Universal Robots URScript: T004_mistralai_Mistral-Large-3-675B-Instruct-2512-NVFP4_edit_perf_rep1.urscript

# Task: T004 — Multi-waypoint SSM pick-place with obstacle avoidance (Optimized)
# Robot: ur5e | Mode: collaborative | Max TCP speed: 0.250 m/s
# Payload: 1.5 kg | Optimized for cycle time

def task_T004():
  TCP_SPEED_CAP = 0.250
  def safe_movel(pose, a, v, r):
    if (v > TCP_SPEED_CAP):
      popup("TCP speed cap exceeded", error=True)
      halt
    end
    movel(pose, a=a, v=v, r=r)
  end

  # [0] Verify E-Stop clear
  if (get_digital_in(0) == True):
    popup("E-Stop active — aborting program.", error=True)
    halt
  end

  # [1] Home position - Increased acceleration
  movej([0.0000, -1.5708, 1.5708, -1.5708, -1.5708, 0.0000], a=2.0000, v=1.0000)

  # [2] WP1 — Above pick station - Increased speed and acceleration
  safe_movel(p[0.400000, -0.250000, 0.350000, 0.0000, 3.1416, 0.0000], 1.2000, 0.2500, 0.0100)

  # [3] WP2 — Descend to pick - Optimized acceleration
  safe_movel(p[0.400000, -0.250000, 0.100000, 0.0000, 3.1416, 0.0000], 1.0000, 0.1000, 0.0)

  # [4] Gripper CLOSE - Parallel execution with next move
  set_digital_out(0, True)
  # [5] Grip settle reduced
  sleep(0.1000)

  # [6] WP3 — Lift above pick - Increased speed and acceleration
  safe_movel(p[0.400000, -0.250000, 0.400000, 0.0000, 3.1416, 0.0000], 1.2000, 0.2500, 0.0150)

  # [7] WP4 — Obstacle avoidance waypoint - Max speed and acceleration
  safe_movel(p[0.250000, 0.000000, 0.400000, 0.0000, 3.1416, 0.0000], 1.5000, 0.2500, 0.0200)

  # [8] WP5 — Above place station - Max speed and acceleration
  safe_movel(p[0.400000, 0.250000, 0.400000, 0.0000, 3.1416, 0.0000], 1.5000, 0.2500, 0.0150)

  # [9] WP6 — Descend to place - Optimized acceleration
  safe_movel(p[0.400000, 0.250000, 0.100000, 0.0000, 3.1416, 0.0000], 1.0000, 0.1000, 0.0)

  # [10] Gripper OPEN - Parallel execution with next move
  set_digital_out(0, False)
  # [11] Release settle reduced
  sleep(0.1000)

  # [12] WP7 — Retract above place - Increased speed and acceleration
  safe_movel(p[0.400000, 0.250000, 0.400000, 0.0000, 3.1416, 0.0000], 1.2000, 0.2500, 0.0100)

  # [13] Return to home - Increased speed and acceleration
  movej([0.0000, -1.5708, 1.5708, -1.5708, -1.5708, 0.0000], a=2.0000, v=1.0000)
end

# Entry point
task_T004()
